(* IEC 61131-3 sources: horner-cscape-mcp/artifacts/projects/Fail_Semicolon_Location_Proj/pous, 1 file *)

(* ---- POU_MissingSemicolon.st ---- *)
PROGRAM POU_MissingSemicolon
VAR
    TargetCount : INT;
END_VAR

TargetCount := 42
END_PROGRAM
